{attribute 'qualified_only'}
{attribute 'strict'}
TYPE E_LimitBasis :
(
	Pcc			:= 0,	// 접속점 기준 (보정 전)
	Device		:= 1	// 설비 기준 (보정 후, PCS 출력 합)
) INT;
END_TYPE

(* stored: Version 1.1.0.1, ProductVersion 3.1.4024.15
   DUT E_LimitBasis: Id {1869ec84-a351-401f-916d-d0d9a42c47df} *)
